(* IEC 61131-3 sources: Versio-VersionControlSystem/fixtures/projects/RefrigeratorControl_FBS/RefrigeratorControl.fbsproj/Device.device.xml.v3^/Plc Logic.plclogic.xml.v3^/Application.application.xml.v3^/Library/Alarm/POUs/FB_Alarm.fb.st^/Protected, 1 file *)

(* ---- _M_Protected.meth.st ---- *)
(* METADATA
{
	"v3Meta": {
		"objectGuid": "523bd15d-dcb8-4ad4-8502-a971302f1b5d"
	}
}
*)
METHOD PROTECTED _M_Protected : BOOL
VAR_INPUT
END_VAR

END_METHOD
